FUNCTION_BLOCK FB_Cylinder
VAR_INPUT
	bExtend		: BOOL;
	nStrokeTicks	: UINT := 5;
END_VAR
VAR_OUTPUT
	bExtended	: BOOL;
END_VAR
VAR
	_nTicks	: UINT;
END_VAR

IF bExtend THEN
	IF _nTicks < nStrokeTicks THEN
		_nTicks := _nTicks + 1;
	END_IF
ELSE
	_nTicks := 0;
END_IF
bExtended := bExtend AND _nTicks >= nStrokeTicks;

METHOD Stroke : UINT
VAR
END_VAR
Stroke := _nTicks;
END_METHOD

END_FUNCTION_BLOCK

(* stored: Version 1.1.0.1, ProductVersion 3.1.4024.12
   POU FB_Cylinder: Id {32a39284-f5a4-49bf-9468-b7abbeb16de3}, SpecialFunc None
   Method Stroke: Id {e9d0598f-e383-4632-a261-a9e833fb80c2} *)
